(* IEC 61131-3 sources: repolevel_ST_code_completion/output/full_case_fixed/repoeval_ProductionLine/readful_result, 4 files *)

(* ---- Motor.st ---- *)
FUNCTION_BLOCK Motor
VAR_INPUT
	MotorI:MotorI;
END_VAR
VAR_OUTPUT
	MotorO:MotorO;
END_VAR
VAR
	WaitTimer: TON;
	InternalSequenceDelay: TIME;
END_VAR

IF MotorI.Overload THEN
	MotorO.FaultStatus := TRUE;
	MotorO.Coil := FALSE;
	RETURN;
END_IF

IF MotorO.FaultStatus = FALSE THEN
WaitTimer.IN := TRUE; // Setting the 'IN' input for the TON block instance.
  WaitTimer.PT := InternalSequenceDelay; // Setting the 'PT' (preset time) input for the TON block instance.
  WaitTimer(); // Executing the TON instance.
END_IF

IF WaitTimer.Q THEN
	MotorO.Coil := TRUE;
WaitTimer.IN := FALSE; // Resetting the 'IN' input for the TON block instance.
  WaitTimer(); // Executing the TON instance to ensure state updates.
END_IF

RETURN;
END_FUNCTION_BLOCK

(* ---- Motor_SetWaitTime.st ---- *)
METHOD SetWaitTime : BOOL
VAR_INPUT
MotorI:MotorI;
SequenceDelay:TIME;
END_VAR
VAR_OUTPUT
MotorO:MotorO;
END_VAR
VAR
WaitTimer:TON;
InternalSequenceDelay:TIME;
END_VAR

InternalSequenceDelay := SequenceDelay;

IF MotorO.FaultStatus = FALSE THEN
// Start the timer when there is no fault
WaitTimer(IN := TRUE, PT := InternalSequenceDelay); // Correctly call TON instance
END_IF

IF WaitTimer.Q THEN
// Activate MotorO coil when WaitTimer indicates timeout
MotorO.Coil := TRUE;
// Stop the timer; no need to check "WaitTimer.IN" explicitly
WaitTimer(IN := FALSE); // Correctly call TON instance again to reset it
END_IF

RETURN;
// Replace incorrect keyword "END_OTHER" with "END_METHOD"
END_METHOD

(* ---- Motor_TurnOff.st ---- *)
METHOD TurnOff : BOOL
VAR_INPUT
	MotorI:MotorI;
END_VAR
VAR_OUTPUT
	MotorO:MotorO;
END_VAR
VAR
	WaitTimer:TON;
	InternalSequenceDelay:TIME;
END_VAR

MotorO.Coil := FALSE;
RETURN;
END_OTHER

(* ---- Motor_TurnOn.st ---- *)
METHOD TurnOn : BOOL
VAR_INPUT
MotorI:MotorI;
END_VAR
VAR_OUTPUT
MotorO:MotorO;
END_VAR
VAR
WaitTimer:TON;
InternalSequenceDelay:TIME;
END_VAR

// Ensure WaitTimer executes only when necessary
IF MotorO.FaultStatus = FALSE THEN
WaitTimer.IN := TRUE;
WaitTimer.PT := InternalSequenceDelay;
WaitTimer(); // Execute the TON function block
END_IF

IF WaitTimer.Q THEN
MotorO.Coil := TRUE;

// Reset the timer only if necessary
IF WaitTimer.IN THEN
 WaitTimer.IN := FALSE;
 WaitTimer(); // Call TON to reflect the reset state
END_IF
END_IF

RETURN;
END_METHOD
